(* IEC 61131-3 sources: daoli-st-library/DL_Algo (part 7) *)

(* ---- FC_DL_SecantIterStep.st ---- *)
(* ============================================================
   DL_Algo / FC_DL_SecantIterStep ｜ v1.0.0 ｜ 2026-11-25
   功能：割线法单步（无导数、四点输入）：x = fX1 − fF1·(fX1−fX0)/(fF1−fF0)，
         并出位移 fDelta；uIter 透传，仅用于差分近零时的扰动方向（偶 +1/奇 −1）
   边界：差分 |fF1−fF0| ≤ 1E-12 → 退化，走相对尺度扰动步 MAX(|x|·1E-3, 1E-6)，
         保证不零步空转；非有限 → 新点/位移写 0（N1），bDegenerate=TRUE
   依赖：仅 IEC 61131-3（ABS / MAX / MOD） ｜ 溯源：DLF-B-ROOTSTEP（内部原创线）
   ============================================================ *)
FUNCTION FC_DL_SecantIterStep : BOOL
VAR_INPUT
    fX0   : LREAL;  // 前一点 [-] / Previous iterate
    fX1   : LREAL;  // 当前点 [-] / Current iterate
    fF0   : LREAL;  // 前一点函数值 [-] / Function value at the previous iterate
    fF1   : LREAL;  // 当前点函数值 [-] / Function value at the current iterate
    uIter : UDINT;  // 迭代序号（透传，仅定扰动方向）[-] / Iteration index passed through
END_VAR
VAR_OUTPUT
    fXnew       : LREAL;  // 割线外推新点 [-] / New secant iterate
    fDelta      : LREAL;  // 本步位移 = fXnew − fX1 [-] / Step displacement
    bDegenerate : BOOL;   // 差分近零或非有限 [-] / Degenerate slope or non-finite value
END_VAR
VAR
    _fDen    : LREAL;  // 差分 = fF1 − fF0 [-] / Difference of function values
    _fJitter : LREAL;  // 退化扰动步长 [-] / Jitter step used when the slope degenerates
END_VAR
VAR CONSTANT
    DL_SEC_EPS   : LREAL := 1.0E-12;  // 差分判零容差 [-] / Slope zero tolerance
    DL_SEC_REL   : LREAL := 1.0E-3;   // 扰动相对尺度系数 [-] / Relative jitter scale
    DL_SEC_FLOOR : LREAL := 1.0E-6;   // 扰动绝对下限 [-] / Absolute jitter floor
END_VAR

(* 段 0：出口预置安全侧（新点 0、位移 0、标退化，N1/N3） *)
FC_DL_SecantIterStep := FALSE;
fXnew := 0.0;  fDelta := 0.0;  bDegenerate := TRUE;

(* 段 1：非有限闸（四个浮点入参全量枚举：NaN 自反，R79/R272） *)
IF (fX0 <> fX0) OR (fX1 <> fX1) OR (fF0 <> fF0) OR (fF1 <> fF1) THEN RETURN; END_IF
(* 段 1b：Inf 双判必须覆盖 fX0/fF0 —— 只判 fX1/fF1 时 fF0=+Inf 使差分 −Inf，
   位移算成 0 却报 bDegenerate=FALSE 且返回 TRUE（静默零步空转） *)
IF ((fX0 - fX0) <> (fX0 - fX0)) OR ((fX1 - fX1) <> (fX1 - fX1))
   OR ((fF0 - fF0) <> (fF0 - fF0)) OR ((fF1 - fF1) <> (fF1 - fF1)) THEN RETURN; END_IF

(* 段 2：差分近零 → 相对尺度扰动（对称试探，防单侧卡死） *)
_fDen := fF1 - fF0;
IF ABS(_fDen) <= DL_SEC_EPS THEN
    _fJitter := MAX(ABS(fX1) * DL_SEC_REL, DL_SEC_FLOOR);
    IF (uIter MOD 2) = 0 THEN
        fXnew := fX1 + _fJitter;              // 偶序号向右
    ELSE
        fXnew := fX1 - _fJitter;              // 奇序号向左
    END_IF
    fDelta := fXnew - fX1;
    bDegenerate := TRUE;  FC_DL_SecantIterStep := TRUE;  RETURN;
END_IF

(* 段 3：割线外推（除子已证 |den| > EPS） *)
fXnew := fX1 - fF1 * (fX1 - fX0) / _fDen;
bDegenerate := FALSE;

(* 段 4：结果复检（非有限回退当前点，出口闸在最后，N4） *)
IF (fXnew <> fXnew) OR ((fXnew - fXnew) <> (fXnew - fXnew)) THEN
    fXnew := fX1;  fDelta := 0.0;  bDegenerate := TRUE;  RETURN;
END_IF
fDelta := fXnew - fX1;
FC_DL_SecantIterStep := TRUE;
END_FUNCTION

(* ---- FC_DL_SettleTimeCalc.st ---- *)
// FC_DL_SettleTimeCalc v1.0.0
// 开源溯源：self-cleanroom / 回路 KPI 族
(*
  道莅工业代码库 | DL_Algo | FC_DL_SettleTimeCalc
  版本: 1.0.0 | 日期: 2026-11-23 | 轮次: R75
  功能: 阶跃响应整定时间：以 ±容差带（相对 y_final）进入判据，扫响应序列
        找最后一次越界采样，整定时间 = 最后越界点之后一拍时刻；
        从未进带 → bSettled=FALSE，带内起步 → 整定时间为 0
  邻件关系: 与 FC_DL_OvershootPctCalc（本批 S22，超调量）成对；与
            FB_DL_WindowExtremaStat（窗口极值统计）差异点：极值件做
            滑窗在线统计，本件为离线序列一次性判据扫描
  序列契约: aResp 为定长显式上界 200 数组，nCount 个有效采样（1..200），
            fTs 为采样周期；本件不改写输入数组
*)
FUNCTION FC_DL_SettleTimeCalc : REAL
VAR_INPUT
    aResp     : ARRAY[1..200] OF REAL;   // 阶跃响应序列（前 nCount 个有效）[工程单位] / Step response samples
    nCount    : INT;                     // 有效采样数 [点]，域 1..200 / Valid sample count, domain 1..200
    fTs       : REAL := 0.1;             // 采样周期 [s]，域 > 0 / Sampling period [s]
    fYFinal   : REAL := 0.0;             // 目标稳态值 [工程单位] / Target steady value
    fBandHalf : REAL := 2.0;             // 容差半带宽 [工程单位]，域 >= 0 / Half tolerance band
END_VAR
VAR_OUTPUT
    bSettled  : BOOL;                    // 序列内已进入容差带并保持 [-] / Settled within band
    bValid    : BOOL;                    // 结果有效回执 [-] / Result validity receipt
    uErrorId  : UDINT;                   // 事件码，0 = 无事件；16#0002_2A01 = 入参域外 / Event code
END_VAR
VAR
    i         : INT;                     // 扫描索引 [点] / Scan index
    nLastViol : INT;                     // 最后越界采样索引 [点]，0 = 从未越界 / Last violating index, 0 = never violated
    fDev      : REAL;                    // 当前偏差 [工程单位] / Current deviation
END_VAR

// —— 段 0：全路径缺省 —— //
bSettled := FALSE;                       // 整定标志预清 / Settled preset
bValid := FALSE;                         // 有效回执预清 / Validity preset
uErrorId := 16#0000;                     // 事件码预清 / Event code preset
nLastViol := 0;                          // 最后越界索引预清（0 = 无越界）/ Last violation preset
FC_DL_SettleTimeCalc := 0.0;             // 返回值缺省零 / Return default zero

// —— 段 1：入参域闸（计数/周期/带宽） —— //
IF (nCount < 1) OR (nCount > 200) OR (fTs <= 0.0) OR (fTs <> fTs)
   OR (fBandHalf < 0.0) OR (fYFinal <> fYFinal) THEN
    uErrorId := 16#0002_2A01;            // 信息级：计数/周期/带宽非法 / Info level: illegal parameters
    RETURN;                              // 不扫描返回 / Return without scan
END_IF

// —— 段 2：序列扫描（找最后一次越出 ±容差带的采样） —— //
FOR i := 1 TO nCount DO                  // 逐点扫描（i ≤ nCount ≤ 200 判界安全）/ Scan points, index safe
    fDev := aResp[i] - fYFinal;          // 与稳态偏差 [工程单位] / Deviation from final
    IF (aResp[i] <> aResp[i]) OR (ABS(fDev) >= 3.0E38) THEN
        uErrorId := 16#0002_2A01;        // 序列含非有限值：拒收（R4 域闸）/ Non-finite sample: reject
        bSettled := FALSE;               // 整定标志回清 / Settled cleared
        RETURN;
    END_IF
    IF ABS(fDev) > fBandHalf THEN        // 越出容差带 / Outside tolerance band
        nLastViol := i;                  // 记录最后越界索引 / Record last violation
    END_IF
END_FOR

// —— 段 3：判据收口（进入带并保持 = 最后越界之后无越界） —— //
IF nLastViol = 0 THEN
    bSettled := TRUE;                    // 全程带内：整定时间 0 / In band from start
    FC_DL_SettleTimeCalc := 0.0;         // 整定时间零 / Settle time zero
ELSE
    IF nLastViol >= nCount THEN
        bSettled := FALSE;               // 末点仍越界：序列内未整定 / Still violating at end
        FC_DL_SettleTimeCalc := 0.0;     // 时间无意义置零 / Time meaningless, zero
    ELSE
        bSettled := TRUE;                // 最后越界后保持带内 / In band after last violation
        FC_DL_SettleTimeCalc := DINT_TO_REAL(nLastViol) * fTs;   // 整定时间 = 越界点后一拍时刻 [s] / Settle time after last violation
    END_IF
END_IF
bValid := TRUE;                          // 有效回执 / Validity receipt
END_FUNCTION

(* ---- FC_DL_SortChuteTimingCalc.st ---- *)
(*
  DL Factory R83 | FC_DL_SortChuteTimingCalc
  功能：按输送速度与到滑槽口距离算分拣释放延时，扣除物件半长与读码延时。
  开源溯源：无（clean-room 自研，依据公开工艺公式，来源=行业通用公式，许可证=MIT，借鉴点=公式结构）
  规则：R1-R21 全遵守
*)
FUNCTION FC_DL_SortChuteTimingCalc : REAL
VAR_INPUT
    fConvSpeedMps : REAL; // 输送线速度 [m/s] / Conveyor speed [m/s]
    fDistM        : REAL; // 读码位到滑槽口距离 [m] / Scanner-to-chute distance [m]
    fItemLenMm    : REAL; // 物件沿输送方向长度 [mm] / Item length along travel [mm]
    fScanDelayMs  : REAL; // 读码与决策固有延时 [ms] / Scan and decision latency [ms]
END_VAR
VAR_OUTPUT
    fReleaseDelayMs : REAL; // 从读码成功到释放的延时 [ms] / Release delay after good read [ms]
    fTransitMs      : REAL; // 纯输送通过时间 [ms] / Pure conveyor transit time [ms]
    fLeadM          : REAL; // 需提前释放的等效距离 [m] / Equivalent lead distance [m]
    xValid          : BOOL; // 计算有效性标志 / Calculation validity flag
END_VAR
// 出口预置：四出口统一预置（R256）
fReleaseDelayMs := 0.0; fTransitMs := 0.0; fLeadM := 0.0; xValid := FALSE;
// 非有限拦截 + 量纲自检 + 速度零闸（R4/R20/R21）
IF NOT (fConvSpeedMps > -1.0E30 AND fConvSpeedMps < 1.0E30) OR NOT (fDistM > -1.0E30 AND fDistM < 1.0E30) OR NOT (fItemLenMm > -1.0E30 AND fItemLenMm < 1.0E30) OR NOT (fScanDelayMs > -1.0E30 AND fScanDelayMs < 1.0E30) OR fConvSpeedMps <= 0.0 OR fDistM < 0.0 OR fItemLenMm < 0.0 OR fScanDelayMs < 0.0 THEN
    FC_DL_SortChuteTimingCalc := -1.0; RETURN;   // 哨兵 -1：非有限或量纲越界 / Sentinel -1
END_IF
// 纯输送时间：m ÷ (m/s) = s，×1000 = ms（分母已判正，量纲自洽）
fTransitMs := (fDistM / fConvSpeedMps) * 1000.0;   // 输送时间 [ms] / Transit time [ms]
// 等效提前距离：物件半长使物件中心先到位，mm ÷ 1000 = m
fLeadM := (fItemLenMm / 1000.0) / 2.0;             // 半长提前量 [m] / Half-length lead [m]
// 释放延时：输送时间 + 读码延时 - 半长对应输送时间（m ÷ m/s × 1000 = ms）
fReleaseDelayMs := fTransitMs + fScanDelayMs - (fLeadM / fConvSpeedMps) * 1000.0; // 释放延时 [ms]
// 物理可实现性闸：延时为负说明读码位过近，判不可分拣
IF fReleaseDelayMs < 0.0 THEN
    fReleaseDelayMs := 0.0;         // 负延时不可执行，钳零 / Negative delay clamped to zero
    xValid          := FALSE;       // 标记不可分拣 / Flag as unsortable
ELSE
    xValid := TRUE;                 // 时序可实现 / Timing feasible
END_IF
FC_DL_SortChuteTimingCalc := fReleaseDelayMs; // 返回释放延时 [ms] / Return release delay [ms]
END_FUNCTION

(* ---- FC_DL_SputterTargetUtilCalc.st ---- *)
(*
  DL Factory R88 | FC_DL_SputterTargetUtilCalc
  功能：按侵蚀环近似算靶材利用率 =已用体积 π(R²-r²)h / 靶体积 πR²t（π 对消），超 80% 提示换靶
  开源溯源：无（clean-room 自研，依据公开工艺公式 靶材利用率体积比定义式，许可证=MIT，借鉴点=公式结构）
  规则：R1-R16 全遵守；R88 简单件标量形（纯标量入参出参，无循环体、无方法、无属性、无数组）
*)
FUNCTION FC_DL_SputterTargetUtilCalc : REAL
VAR_INPUT
    fTargetRmm : REAL := 150.0; // 靶材有效半径 R [mm] / target radius [mm]
    fErosionRmm : REAL := 80.0; // 侵蚀环内边界半径 r（环宽 R-r） [mm] / erosion ring inner radius [mm]
    fErosionDepthMm : REAL := 4.0; // 侵蚀环最大深度 h [mm] / erosion depth [mm]
    fTargetThkMm : REAL := 10.0; // 靶材原始厚度 t [mm] / original target thickness [mm]
    fReplacePct : REAL := 80.0; // 换靶提示阈值（利用率超过即换靶） [%] / replacement threshold [%]
END_VAR
VAR_OUTPUT
    fUtilPct : REAL; // 靶材利用率（体积比） [%] / target utilisation [%]
    xReplace : BOOL; // TRUE=利用率超过阈值，需换靶 [-] / TRUE when replacement is due [-]
END_VAR
VAR
    fTargetVolMm3 : REAL; // 靶材总体积 πR²t（除零判据） [mm³] / total target volume, the divisor [mm^3]
    fR2MinusR2 : REAL; // R²-r²（符号闸判据） [mm²] / difference of squares [mm^2]
END_VAR

// 段 1｜出口预置
FC_DL_SputterTargetUtilCalc := -1.0; // 哨兵返回 -1（无效） [-] / sentinel return -1, invalid [-]
fUtilPct := 0.0; // 利用率预置零 [%] / utilisation preset zero [%]
xReplace := FALSE; // 换靶位预置 FALSE（未判定前不提示） [-] / replace flag preset false [-]

// 段 2｜非有限拦截 + 域闸
IF NOT (fTargetRmm > -1.0E30 AND fTargetRmm < 1.0E30) OR NOT (fErosionRmm > -1.0E30 AND fErosionRmm < 1.0E30) OR NOT (fErosionDepthMm > -1.0E30 AND fErosionDepthMm < 1.0E30) THEN
    RETURN; // 靶半径/侵蚀半径/侵蚀深度任一非有限即拒算 [-] / any non finite input rejected [-]
END_IF
IF NOT (fTargetThkMm > -1.0E30 AND fTargetThkMm < 1.0E30) OR NOT (fReplacePct > -1.0E30 AND fReplacePct < 1.0E30) THEN
    RETURN; // 靶厚/换靶阈值任一非有限则判据静默失效，故先拦 [-] / these pins must be finite [-]
END_IF
IF fTargetRmm < 1.0E-9 OR fTargetThkMm < 1.0E-9 OR fErosionDepthMm < 0.0 THEN
    RETURN; // 靶半径/靶厚正域闸（分母）+ 侵蚀深度非负闸 [mm] / positive geometry gates [mm]
END_IF
IF fErosionRmm < 0.0 OR fErosionRmm >= fTargetRmm THEN
    RETURN; // 侵蚀环几何闸：0≤r<R，否则环带面积为零或负 [mm] / erosion ring geometry gate [mm]
END_IF
IF fReplacePct <= 0.0 OR fReplacePct > 100.0 THEN
    RETURN; // 换靶阈值区间闸 (0,100]：超出则判据无意义 [%] / replacement threshold gate [%]
END_IF

// 段 3｜计算（侵蚀环按矩形截面近似，π 在比值中约去）
fR2MinusR2 := fTargetRmm * fTargetRmm - fErosionRmm * fErosionRmm; // mm² - mm² = mm²，环带相当面积 [mm²] / [mm^2]
fTargetVolMm3 := 3.14159265 * fTargetRmm * fTargetRmm * fTargetThkMm; // 无量纲 × mm² × mm = mm³，靶体积 [mm³] / [mm^3]
IF fR2MinusR2 <= 0.0 OR fTargetVolMm3 < 1.0E-9 THEN
    RETURN; // 平方差闸 + 除法前分母闸：两者须为正，否则体积链失效 [mm², mm³] / volume chain gates
END_IF
fUtilPct := 3.14159265 * fR2MinusR2 * fErosionDepthMm / fTargetVolMm3 * 100.0; // (mm³ ÷ mm³) × 100 = %，体积利用率 [%] / [%]

// 段 4｜判定与饱和
IF NOT (fUtilPct > -1.0E30 AND fUtilPct < 1.0E30) THEN
    RETURN; // 结果非有限再拦一次 [-] / re-check the result for finiteness [-]
END_IF
IF fUtilPct > 100.0 THEN
    fUtilPct := 100.0; // 上饱和：体积比不可能超过 100%，超出按 100% 夹紧 [%] / saturate at 100 percent [%]
END_IF
xReplace := fUtilPct > fReplacePct; // 严格大于阈值为需换靶，等于阈值仍可继续 [%] / strict compare [%]

// 段 5｜出口自检
IF fUtilPct < 0.0 THEN
    RETURN; // 出口自检：利用率不得为负（负值说明几何参数错） [%] / utilisation must not be negative [%]
END_IF
FC_DL_SputterTargetUtilCalc := fUtilPct; // 返回靶材利用率 [%] / return the target utilisation [%]
END_FUNCTION

(* ---- FC_DL_SurfaceRoughnessRzFromRaCalc.st ---- *)
(*
  DL Factory R88 | FC_DL_SurfaceRoughnessRzFromRaCalc
  功能：由 Ra 按经验因子换算 Rz（Rz≈k·Ra，车/磨区间 k=3.5~5.0），并判定因子是否落在经验带内
  开源溯源：无（clean-room 自研，依据公开工艺公式 Ra-Rz 经验换算式 Rz≈(3.5~5.0)·Ra，许可证=MIT，借鉴点=公式结构）
  规则：R1-R16 全遵守；R88 简单件标量形（纯标量入参出参，无循环体、无方法、无属性、无数组）
*)
FUNCTION FC_DL_SurfaceRoughnessRzFromRaCalc : REAL
VAR_INPUT
    fRaUm : REAL := 1.6; // 算术平均偏差 Ra [µm] / arithmetic mean roughness Ra [um]
    fProcessFactor : REAL := 4.0; // 工艺经验因子 k（车/磨 3.5~5.0，非标准定义） [-] / empirical process factor [-]
    fMinFactor : REAL := 3.5; // 经验带下限 [-] / lower empirical band [-]
    fMaxFactor : REAL := 5.0; // 经验带上限 [-] / upper empirical band [-]
END_VAR
VAR_OUTPUT
    fRzUm : REAL; // 十点高度 Rz 估计值 [µm] / estimated Rz [um]
    xInBand : BOOL; // TRUE=所用因子落在经验带内，估计可信 [-] / TRUE when the factor is inside the band [-]
END_VAR
VAR
    fFactorLo : REAL; // 实际参与计算的因子下限（缓存） [-] / lower factor bound in use [-]
    fFactorHi : REAL; // 实际参与计算的因子上限（缓存） [-] / upper factor bound in use [-]
END_VAR

// 段 1｜出口预置
FC_DL_SurfaceRoughnessRzFromRaCalc := -1.0; // 哨兵返回 -1（无效） [-] / sentinel return -1, invalid [-]
fRzUm := 0.0; // Rz 估计值预置零 [µm] / Rz estimate preset zero [um]
xInBand := FALSE; // 带宽位预置 FALSE（未判定前不认可信） [-] / band flag preset false [-]
fFactorLo := 0.0; // 因子下限缓存预置零 [-] / lower factor preset zero [-]
fFactorHi := 0.0; // 因子上限缓存预置零 [-] / upper factor preset zero [-]

// 段 2｜非有限拦截 + 域闸
IF NOT (fRaUm > -1.0E30 AND fRaUm < 1.0E30) OR NOT (fProcessFactor > -1.0E30 AND fProcessFactor < 1.0E30) THEN
    RETURN; // Ra/工艺因子任一非有限即拒算 [-] / any non finite input rejected [-]
END_IF
IF NOT (fMinFactor > -1.0E30 AND fMinFactor < 1.0E30) OR NOT (fMaxFactor > -1.0E30 AND fMaxFactor < 1.0E30) THEN
    RETURN; // 经验带上下限任一非有限则判据静默失效，故先拦 [-] / band limits must be finite [-]
END_IF
IF fRaUm < 0.0 THEN
    RETURN; // Ra 非负闸：粗糙度不得为负 [µm] / non negative Ra gate [um]
END_IF
IF fProcessFactor < 1.0 OR fProcessFactor > 10.0 THEN
    RETURN; // 因子工程域闸 (1,10)：越界则换算关系不再成立 [-] / factor domain gate [-]
END_IF
IF fMinFactor <= 0.0 OR fMaxFactor <= fMinFactor THEN
    RETURN; // 经验带自洽闸：下限须为正、上限须严格大于下限 [-] / band consistency gate [-]
END_IF

// 段 3｜计算（经验换算，不是标准定义：Rz 与 Ra 无通用解析关系）
fFactorLo := fMinFactor; // 取经验带下限参与判定 [-] / take the lower factor bound [-]
fFactorHi := fMaxFactor; // 取经验带上限参与判定 [-] / take the upper factor bound [-]
fRzUm := fProcessFactor * fRaUm; // 无量纲 × µm = µm，Rz≈k·Ra [µm] / [-] x [um] = [um]

// 段 4｜判定与饱和
IF NOT (fRzUm > -1.0E30 AND fRzUm < 1.0E30) THEN
    RETURN; // 结果非有限再拦一次（防溢出成 Inf） [µm] / re-check the result for finiteness [um]
END_IF
xInBand := (fProcessFactor >= fFactorLo) AND (fProcessFactor <= fFactorHi); // 因子与经验带双侧直比 [-] / factor against the empirical band [-]

// 段 5｜出口自检
IF fRzUm < fRaUm THEN
    RETURN; // 出口自检：Rz 不应小于 Ra（因子域闸已保证 k>1，否则换算链被破坏） [µm] / Rz must not fall below Ra [um]
END_IF
FC_DL_SurfaceRoughnessRzFromRaCalc := fRzUm; // 返回 Rz 估计值 [µm] / return the estimated Rz [um]
END_FUNCTION

(* ---- FC_DL_TcToFilterCoeff.st ---- *)
//==============================================================================
// 函数：FC_DL_TcToFilterCoeff ｜ 中文名称：时间常数→离散一阶滤波系数换算原子
// 所属子库：DL_Algo ｜ 版本：v1.0.0 ｜ 日期：2026-11-23
// 兼容：CODESYS V3.5+ / TwinCAT 3 / 汇川 InoProShop（纯标准库）
// 功能描述：α = Ts/(Ts + Tc) 离散一阶低通滤波系数换算原子（后向欧拉口径）。
//           分工声明：系数原子属本件；一阶滤波本体（驻留状态、逐拍迭代）
//           属 FB_DL_LowPassFilter，互不替代——该件头注释与本件互引，
//           上层先经本件换算 α 再注入滤波本体。
// 开源溯源 (Origin)：原创实现（自研-std 标准包装线，零外部源码行，clean-room
//           独立编写）
// 公开接口清单：输入 fTs / fTc；输出 返回值 / bValid
// 单位表：fTs / fTc [秒] / 返回值 α [1]（无量纲系数）
// 输入契约：fTs 须与实际任务周期一致（任务周期变更须重算重注入）；fTc >= 0
//           合法（0 = 直通旁路口径）。
// 输出契约：返回值为后向欧拉离散滤波系数，域 (0, 1]；bValid = FALSE 拍
//           返回哨兵 0.0，禁注入 FB_DL_LowPassFilter。
// 错误码表：纯函数无状态机码轨；无效输入经 bValid = FALSE 表达（哨兵返回
//           0.0），本件不占用 16#0002 段码位（邻件免让位）
// 状态机：N/A（纯函数，无状态，可重入）
// 边界行为：① fTs <= 0（采样周期非法）→ 拒绝（bValid := FALSE，哨兵 0.0）；
//           ② fTc < 0（时间常数非法）→ 拒绝；fTc = 0 合法（α = 1 直通）；
//           ③ 分母 (Ts + Tc) 先过正域闸再除（防除零强制闸）；
//           ④ 非有限输入 → 哨兵 0.0 返回；
//           ⑤ α 输出域 (0, 1]，数学上由分子分母同号保证，仍出口钳位兜底。
// 修订历史：v1.0.0 2026-11-23 首版（R73 派单 · 批 3 · 序 17）
//==============================================================================

(*------------------------------------------------------------------------------
 * 调用示例：fA := FC_DL_TcToFilterCoeff(fTs := 0.01, fTc := 0.5,
 *                                       bValid => bOk);
 * 注意：α = 0.01/0.51 ≈ 0.0196；α 注入 FB_DL_LowPassFilter 前必须 bOk。
 * 组装说明：① 与 FB_DL_LowPassFilter 互引分工：本件出系数、该件做逐拍
 *             滤波本体，bValid = FALSE 拍 α 不得注入滤波本体；
 *           ② fTs 应与实际任务周期一致（任务周期变更须重算并重注入）；
 *           ③ fTc = 0 时 α = 1 直通（滤波旁路口径，上层据此可做旁路）。
 *-----------------------------------------------------------------------------*)
FUNCTION FC_DL_TcToFilterCoeff : LREAL
VAR_INPUT
    fTs     : LREAL;                   // 采样周期 [秒]，有效域 (0, +∞) / Sampling period [s]
    fTc     : LREAL;                   // 滤波时间常数 [秒]，有效域 [0, +∞) / Filter time constant [s]
END_VAR
VAR_OUTPUT
    bValid  : BOOL;                    // 结果有效标志，FALSE 时返回哨兵 0.0 / Result validity flag
END_VAR
VAR CONSTANT
    DL_TC_EPS  : LREAL := 1.0E-12;     // 分母正域闸容差 [秒] / Denominator gate tolerance [s]
    DL_TC_INF  : LREAL := 1.7976931348623157E308; // LREAL 幅值上限 / LREAL magnitude ceiling
    DL_TC_ZERO : LREAL := 0.0;         // 无效哨兵返回值 / Sentinel return for invalid
    DL_TC_ONE  : LREAL := 1.0;         // α 上界（直通口径）/ Alpha ceiling, pass-through
END_VAR

// ---- 段 1｜出口默认值（纯函数无实例，无定时器/沿刷新义务）----
bValid := FALSE;                      // 缺省无效 / Invalid by default

// ---- 段 2｜输入防御：非有限值（NaN 自反判 + Inf 幅值判，R79）----
IF (fTs <> fTs) OR (ABS(fTs) > DL_TC_INF)
   OR (fTc <> fTc) OR (ABS(fTc) > DL_TC_INF) THEN
    FC_DL_TcToFilterCoeff := DL_TC_ZERO; // 无效输入：哨兵零返回 / Invalid input, sentinel zero return
    RETURN;                            // 结构早退 / early exit
END_IF

// ---- 段 3｜域闸：Ts 正域 + Tc 非负域（fTc = 0 合法 = α 直通）----
IF (fTs <= DL_TC_EPS) OR (fTc < 0.0) THEN
    FC_DL_TcToFilterCoeff := DL_TC_ZERO; // 域外拒绝：哨兵零返回 / Out of domain, refused
    RETURN;                            // 结构早退 / early exit
END_IF

// ---- 段 4｜换算主体：α = Ts/(Ts + Tc)，分母先过正域闸（防除零强制闸）----
IF (fTs + fTc) <= DL_TC_EPS THEN
    FC_DL_TcToFilterCoeff := DL_TC_ZERO; // 分母退化拒绝（理论上不可达，仍强制闸）/ Degenerate denominator, gated
    RETURN;                            // 结构早退 / early exit
END_IF
FC_DL_TcToFilterCoeff := fTs / (fTs + fTc); // 滤波系数 [1] / Filter coefficient [1]
IF FC_DL_TcToFilterCoeff > DL_TC_ONE THEN
    FC_DL_TcToFilterCoeff := DL_TC_ONE; // α 上界钳位兜底（浮点噪声防护）/ Alpha ceiling clamp
END_IF
bValid := TRUE;                       // 全部防御通过：结果有效 / Result valid
END_FUNCTION

(* ---- FC_DL_TernaryNarrowIterStep.st ---- *)
(* ============================================================
   DL_Algo / FC_DL_TernaryNarrowIterStep ｜ v1.0.0 ｜ 2026-11-25
   功能：三分法单步（三点等分比较后收缩）。探针 m1 = a + L/3、m2 = b − L/3，
         其函数值由调用方求值后回灌：fF1<fF2 → 保 [a,m2]；fF1>fF2 → 保 [m1,b]；
         两者容差判等 → 保 [m1,m2]。出新区间与实测收缩比（2/3 或 1/3）
   边界：长度 ≤ 1E-12 → 区间不收缩、fRatio=1（不虚报）；函数值非有限 →
         原区间回传、fRatio=1、返回 FALSE（N1：判据与实值同源）
   依赖：仅 IEC 61131-3（ABS / MIN / MAX） ｜ 溯源：DLF-B-ROOTSTEP（内部原创线）
   ============================================================ *)
FUNCTION FC_DL_TernaryNarrowIterStep : BOOL
VAR_INPUT
    fA  : LREAL;  // 区间下界 [-] / Lower interval bound
    fB  : LREAL;  // 区间上界 [-] / Upper interval bound
    fF1 : LREAL;  // 左三分点 m1 处函数值 [-] / Function value at the left trisection point
    fF2 : LREAL;  // 右三分点 m2 处函数值 [-] / Function value at the right trisection point
END_VAR
VAR_OUTPUT
    fAnew  : LREAL;  // 新区间下界 [-] / New lower bound
    fBnew  : LREAL;  // 新区间上界 [-] / New upper bound
    fRatio : LREAL;  // 实测收缩比 = 新宽/原宽 [-] / Measured shrink ratio
END_VAR
VAR
    _fLen : LREAL;  // 原区间长度 [-] / Original interval length
    _fM1  : LREAL;  // 左三等分点 [-] / Left trisection point
    _fM2  : LREAL;  // 右三等分点 [-] / Right trisection point
    _fLo  : LREAL;  // 区间小端 [-] / Smaller interval end
    _fHi  : LREAL;  // 区间大端 [-] / Larger interval end
END_VAR
VAR CONSTANT
    DL_TNY_EPS : LREAL := 1.0E-12;  // 函数值判等容差与长度判零 [-] / Equality tolerance and length floor
END_VAR

(* 段 0：出口预置安全侧（新区间=原区间、收缩比 1，N3） *)
FC_DL_TernaryNarrowIterStep := FALSE;
fAnew := 0.0;  fBnew := 0.0;  fRatio := 1.0;

(* 段 1：非有限闸 *)
IF (fA <> fA) OR (fB <> fB) OR (fF1 <> fF1) OR (fF2 <> fF2) THEN RETURN; END_IF
IF ((fB - fA) - (fB - fA)) <> ((fB - fA) - (fB - fA)) THEN RETURN; END_IF

(* 段 2：闸后原样回传（fRatio=1 表示本步未收缩）与长度退化闸 *)
fAnew := fA;  fBnew := fB;  fRatio := 1.0;
_fLo := MIN(fA, fB);  _fHi := MAX(fA, fB);
_fLen := _fHi - _fLo;
IF _fLen <= DL_TNY_EPS THEN
    fAnew := _fLo;  fBnew := _fHi;  fRatio := 1.0;
    FC_DL_TernaryNarrowIterStep := TRUE;  RETURN;
END_IF

(* 段 3：三等分两点与三点比较收缩（判等带容差，方向分列） *)
_fM1 := _fLo + _fLen / 3.0;
_fM2 := _fHi - _fLen / 3.0;
IF ABS(fF1 - fF2) <= DL_TNY_EPS THEN
    fAnew := _fM1;  fBnew := _fM2;            // 两侧等高：保中间三分之一
ELSIF fF1 < fF2 THEN
    fAnew := _fLo;  fBnew := _fM2;            // 左低：保左侧三分之二
ELSE
    fAnew := _fM1;  fBnew := _fHi;            // 右低：保右侧三分之二
END_IF

(* 段 4：实测收缩比 + 越域回退（出口与判据同源，N4） *)
fRatio := (fBnew - fAnew) / _fLen;            // 除子已证 > EPS
IF (fRatio <> fRatio) OR (fRatio < 0.0) OR (fRatio > 1.0) THEN
    fAnew := _fLo;  fBnew := _fHi;  fRatio := 1.0;  RETURN;
END_IF
FC_DL_TernaryNarrowIterStep := TRUE;
END_FUNCTION

(* ---- FC_DL_VacuumPumpdownTimeCalc.st ---- *)
(*
  DL Factory R88 | FC_DL_VacuumPumpdownTimeCalc
  功能：算抽气时间 t=(V/S)·ln(p0/p)，压力比须大于 1 才有效，超 600 s 提示抽速不足
  开源溯源：无（clean-room 自研，依据公开工艺公式 粗抽时间式 t=(V/S)·ln(p0/p)，许可证=MIT，借鉴点=公式结构）
  规则：R1-R16 全遵守；R88 简单件标量形（纯标量入参出参，无循环体、无方法、无属性、无数组）
*)
FUNCTION FC_DL_VacuumPumpdownTimeCalc : REAL
VAR_INPUT
    fVolL : REAL := 100.0; // 腔室容积 V [L] / chamber volume [L]
    fPumpSpeedLps : REAL := 10.0; // 泵有效抽速 S（工作压力段平均值） [L/s] / effective pumping speed [L/s]
    fPStartPa : REAL := 101325.0; // 起始压力 p0 [Pa] / starting pressure [Pa]
    fPEndPa : REAL := 1.0; // 目标压力 p [Pa] / target pressure [Pa]
    fLimitS : REAL := 600.0; // 抽气时间上限 [s] / pumpdown time limit [s]
END_VAR
VAR_OUTPUT
    fTimeS : REAL; // 抽气时间 t [s] / pumpdown time [s]
    xTooLong : BOOL; // TRUE=抽气时间超过上限，抽速不足 [-] / TRUE when the time exceeds the limit [-]
END_VAR
VAR
    fRatio : REAL; // 压力比 p0/p（LN 自变量，须 >1） [-] / pressure ratio, the LN argument [-]
    fVolPerSpeedS : REAL; // V/S 时间常数（除零判据） [s] / time constant, the divisor [s]
END_VAR

// 段 1｜出口预置
FC_DL_VacuumPumpdownTimeCalc := -1.0; // 哨兵返回 -1（无效） [-] / sentinel return -1, invalid [-]
fTimeS := 0.0; // 抽气时间预置零 [s] / pumpdown time preset zero [s]
xTooLong := FALSE; // 过久位预置 FALSE（未判定前不报警） [-] / too-long flag preset false [-]

// 段 2｜非有限拦截 + 域闸
IF NOT (fVolL > -1.0E30 AND fVolL < 1.0E30) OR NOT (fPumpSpeedLps > -1.0E30 AND fPumpSpeedLps < 1.0E30) OR NOT (fLimitS > -1.0E30 AND fLimitS < 1.0E30) THEN
    RETURN; // 容积/抽速/时间上限任一非有限即拒算 [-] / any non finite input rejected [-]
END_IF
IF NOT (fPStartPa > -1.0E30 AND fPStartPa < 1.0E30) OR NOT (fPEndPa > -1.0E30 AND fPEndPa < 1.0E30) THEN
    RETURN; // 起始/目标压力任一非有限即拒算 [Pa] / any non finite pressure rejected [Pa]
END_IF
IF fVolL < 1.0E-9 OR fPumpSpeedLps < 1.0E-9 OR fLimitS <= 0.0 THEN
    RETURN; // 容积与抽速正域闸（分母）+ 时间上限正域闸 [L, L/s, s] / positive gates
END_IF
IF fPStartPa < 1.0E-9 OR fPEndPa < 1.0E-9 OR fPStartPa <= fPEndPa THEN
    RETURN; // 压力正域闸（LN 自变量）+ 压力比闸：p0 须大于 p，否则 LN≤0 [Pa] / pressure ratio gate [Pa]
END_IF

// 段 3｜计算
fVolPerSpeedS := fVolL / fPumpSpeedLps; // L ÷ (L/s) = s，时间常数 V/S [s] / [s]
IF fVolPerSpeedS < 1.0E-9 THEN
    RETURN; // 除法后复核：时间常数须为正，否则结果失去物理意义 [s] / the constant must stay positive [s]
END_IF
fRatio := fPStartPa / fPEndPa; // Pa ÷ Pa = 无量纲，压力比 [-] / dimensionless ratio [-]
IF fRatio <= 1.0 THEN
    RETURN; // LN 自变量闸：比值必须大于 1，否则对数为非正 [-] / the LN argument must exceed one [-]
END_IF
fTimeS := fVolPerSpeedS * LN(fRatio); // s × 无量纲 = s，抽气时间 [s] / [s] x [-] = [s]

// 段 4｜判定与饱和
IF NOT (fTimeS > -1.0E30 AND fTimeS < 1.0E30) THEN
    RETURN; // 结果非有限再拦一次 [-] / re-check the result for finiteness [-]
END_IF
xTooLong := fTimeS > fLimitS; // 严格大于上限为过久，等于上限仍判合格 [s] / strict compare [s]

// 段 5｜出口自检
IF fTimeS < 0.0 THEN
    RETURN; // 出口自检：抽气时间不得为负（负值说明压力比给反） [s] / time must not be negative [s]
END_IF
FC_DL_VacuumPumpdownTimeCalc := fTimeS; // 返回抽气时间 [s] / return the pumpdown time [s]
END_FUNCTION

(* ---- FC_DL_VaporPressureSat.st ---- *)
//==============================================================================
// 函数：FC_DL_VaporPressureSat ｜ 中文名称：饱和水蒸气压计算（焓湿图族公式基准原子）
// 所属子库：DL_Algo ｜ 版本：v1.0.0 ｜ 兼容：CODESYS V3.5+ / TwinCAT 3 / 汇川 InoProShop
// 功能描述：Magnus-Tetens（过水面参数化）饱和水蒸气压计算，焓湿图全参族
//           （含湿量/湿球/露点逆运算/混风点）的饱和压唯一属主件，族内其余
//           四件一律调用本件取饱和压，禁止各自内联公式（常量单源，防口径
//           漂移）；与 FC_DL_DewPointCalc 系数口径一致（a=17.625、b=243.04、
//           E0=610.94 Pa），属主转移声明：露点族饱和压口径自本件起收口。
// 开源溯源 (Origin)：改写自 OSCAT Building 行为定义（OSCAT 许可，仅行为定义，零代码行）——道莅 clean-room 实现
// 单位表：T[°C] / p_ws[Pa]
// 错误码表：16#0002_2D01 信息级（温度域外已钳位照算，不置 bError）/ 16#0002_2D10
//           故障级（输入非有限或结果溢出，置 bError）/ 16#0002_2D02、16#0002_2D11、
//           16#0002_2D12 预留禁用（不得挪用）
// 状态机：N/A（纯函数，无状态；同输入必得同输出）
// 边界行为：① 温度域外（-40~100 °C 外）钳位照算 + 信息 2D01 + bClamped，
//           低温干燥是合法工况，不置故障；② 非有限输入（NaN/±Inf）→ 故障
//           2D10、bValid := FALSE、fPvSat := 0、返回 FALSE；③ EXP 上溢拦
//           （结果幅值 > 1.7976931348623157E308 复检）→ 故障 2D10 复用
//           （R90 不加码：同属"数值结果不可用"一类，头注释留档复用理由）；
//           异常路径输出为确定值 0，绝不输出未初始化值。
// 修订历史：v1.0.0 2026-11-17 首版（R23 派单 · T1-2 焓湿图族拆分① · 全族公式基准）
//==============================================================================

(*------------------------------------------------------------------------------
 * 调用示例：bOk := FC_DL_VaporPressureSat(fTempC := 25.0, fPvSat => fPws,
 *                                         bClamped => bC, eErr => uE);
 * 族内引用：FC_DL_HumidityRatioCalc / FC_DL_WetBulbTempCalc /
 *           FC_DL_RhFromDewPoint / FC_DL_MixAirStateCalc 一律经本件取饱和压。
 *-----------------------------------------------------------------------------*)
FUNCTION FC_DL_VaporPressureSat : BOOL
VAR_INPUT
    fTempC    : LREAL;                   // 空气温度 [摄氏度]，有效域 -40.0..100.0，域外钳位照算 / Air temperature [degC], valid range -40.0..100.0, clamped outside
END_VAR
VAR_OUTPUT
    fPvSat    : LREAL;                   // 饱和水蒸气压 [Pa] / Saturation vapor pressure [Pa]
    bClamped  : BOOL;                    // TRUE = 输入已钳位，结果按趋势参考 / TRUE = input clamped, result for trend reference only
    eErr      : UDINT;                   // 错误码，0 = 无错 / Error code, 0 = no error
    bError    : BOOL;                    // 故障级标志，仅故障级错误置位 / Fault-class flag, set only on fault-level codes
    bValid    : BOOL;                    // 输出可用标志 / Outputs usable flag
END_VAR
VAR CONSTANT
    DL_PSV_TMIN  : LREAL := -40.0;       // Magnus-Tetens 有效域下限 [摄氏度] / Magnus-Tetens valid range low [degC]
    DL_PSV_TMAX  : LREAL := 100.0;       // Magnus-Tetens 有效域上限 [摄氏度] / Magnus-Tetens valid range high [degC]
    DL_PSV_E0    : LREAL := 610.94;      // 0 摄氏度饱和水汽压基准 [Pa] / Reference saturation pressure at 0 degC [Pa]
    DL_PSV_A     : LREAL := 17.625;      // Magnus 系数 a [1]，与 FC_DL_DewPointCalc 同口径 / Magnus coefficient a [1], same as dew point FC
    DL_PSV_B     : LREAL := 243.04;      // Magnus 系数 b [摄氏度] / Magnus coefficient b [degC]
    DL_PSV_EPS   : LREAL := 1.0E-6;      // 浮点判零容差 / Float zero tolerance
    DL_PSV_INF   : LREAL := 1.7976931348623157E308; // LREAL 幅值上限，EXP 上溢复检基准 / LREAL magnitude ceiling, EXP overflow recheck bound
END_VAR
VAR
    fTEff   : LREAL;                     // 钳位后的生效温度 [摄氏度] / Effective clamped temperature [degC]
    fDenom  : LREAL;                     // Magnus 分母 (b+T) [摄氏度] / Magnus denominator (b+T) [degC]
    fResult : LREAL;                     // 公式原始结果 [Pa]，有限性复检前暂存 / Raw formula result [Pa], staged before the finiteness recheck
END_VAR

(*------------------------------------------------------------------------------
 * 段 1｜出口默认值：入口即赋确定值，任何提前 RETURN 前输出已确定
 *      Exit defaults: outputs assigned deterministically on entry
 *-----------------------------------------------------------------------------*)
FC_DL_VaporPressureSat := FALSE;         // 返回值默认无效 / Return value preset invalid
fPvSat := 0.0;                           // 饱和压默认置零 / Saturation pressure preset to zero
bClamped := FALSE;                       // 钳位标志默认 FALSE / Clamped flag preset FALSE
eErr := 16#0000_0000;                    // 错误码先清零 / Error code cleared first
bError := FALSE;                         // 故障标志先清零 / Fault flag cleared first
bValid := FALSE;                         // 可用标志先清零 / Usable flag cleared first

(*------------------------------------------------------------------------------
 * 段 2｜非有限值防御：NaN 用 (x<>x) 判，Inf 用双侧幅值判（R79 口径）
 *      Non-finite defense: NaN via (x<>x), Inf via two-sided magnitude bound
 *-----------------------------------------------------------------------------*)
IF (fTempC <> fTempC) OR (fTempC < -DL_PSV_INF) OR (fTempC > DL_PSV_INF) THEN
    eErr   := 16#0002_2D10;              // 故障级：输入非有限（NaN/Inf） / Fault: non-finite input
    bError := TRUE;                      // 故障级码位必须同时置故障标志（R45 配对） / Fault code paired with the fault flag
    bValid := FALSE;                     // 输出不可用 / Outputs unusable
    RETURN;                              // 异常路径出口，fPvSat 保持确定值 0 / Error path exit, output stays deterministic zero
END_IF

(*------------------------------------------------------------------------------
 * 段 3｜温度钳位：域外按趋势参考照算，信息级不置故障（低温干燥合法工况）
 *      Temperature clamping: out-of-domain treated as trend reference, info only
 *-----------------------------------------------------------------------------*)
IF (fTempC < DL_PSV_TMIN) OR (fTempC > DL_PSV_TMAX) THEN
    fTEff := MIN(MAX(fTempC, DL_PSV_TMIN), DL_PSV_TMAX); // 双侧钳位到有效域 / Two-sided clamp into valid range
    bClamped := TRUE;                    // 钳位声明置位 / Clamped flag raised
    eErr := 16#0002_2D01;                // 信息级：温度已钳位（不置 bError） / Info: temperature clamped, no fault flag
ELSE
    fTEff := fTempC;                     // 合法温度原值生效 / Valid temperature applied as-is
END_IF

(*------------------------------------------------------------------------------
 * 段 4｜Magnus-Tetens 主体：p_ws = 610.94·EXP(17.625·T/(T+243.04))
 *      分母 (b+T) 由 T >= -40 保证恒正，仍做防御性双检（防除零）
 *      Magnus-Tetens core, denominator guarded even though always positive
 *-----------------------------------------------------------------------------*)
fDenom := DL_PSV_B + fTEff;              // Magnus 分母 [摄氏度] / Magnus denominator [degC]
IF ABS(fDenom) <= DL_PSV_EPS THEN
    eErr   := 16#0002_2D10;              // 故障级：分母退化复用非有限码（R90） / Fault: degenerate denominator, code reused
    bError := TRUE;                      // 置故障标志 / Raise the fault flag
    bValid := FALSE;                     // 输出不可用 / Outputs unusable
    RETURN;
END_IF
fResult := DL_PSV_E0 * EXP(DL_PSV_A * fTEff / fDenom); // 饱和水蒸气压原始结果 [Pa] / Raw saturation vapor pressure [Pa]

(*------------------------------------------------------------------------------
 * 段 5｜结果有限性复检：EXP 上溢拦（R90 复用 2D10，理由：同属数值结果
 *      不可用一类，不新开码位）
 *      Result finiteness recheck, EXP overflow folded into 2D10 per R90
 *-----------------------------------------------------------------------------*)
IF (fResult <> fResult) OR (fResult > DL_PSV_INF) OR (fResult < -DL_PSV_INF) THEN
    fPvSat := 0.0;                       // 溢出结果丢弃，输出确定值 0 / Overflowed result discarded, output zero
    eErr   := 16#0002_2D10;              // 故障级：结果溢出复用（R90） / Fault: result overflow, code reused
    bError := TRUE;                      // 置故障标志 / Raise the fault flag
    bValid := FALSE;                     // 输出不可用 / Outputs unusable
    RETURN;
END_IF

fPvSat := fResult;                       // 有限结果出口 / Finite result outlet
bValid := TRUE;                          // 输出可用 / Outputs usable
FC_DL_VaporPressureSat := TRUE;          // 返回 TRUE = 计算有效 / Return TRUE = computation valid
END_FUNCTION

(* ---- FC_DL_WaterEnthalpy.st ---- *)
(*==============================================================================
 * 组件名称 (Component)  : FC_DL_WaterEnthalpy
 * 所属子库 (Sublibrary) : DL_Algo
 * 当前版本 (Version)    : 1.0.0
 * 兼容性   (Platform)   : CODESYS 3.5 / TwinCAT 3 / 汇川 InoProShop / Machine Expert
 *                         仅依赖 Standard.library（ABS），零厂商方言
 * 功能描述 (Function)   : 0~150 摄氏度液态水的比焓，以 0 摄氏度饱和液水为焓基准，
 *                         同时给出「0 摄氏度到当前温度的平均比热」。
 *                         现场用途：冷热量表按质量流量乘比焓差结算、板换换热量核算、
 *                         锅炉给水与回水焓差、蓄冷水罐冷量统计。
 *                         用固定 4.186 千焦每千克开尔文替代真实比焓，在 70~90 摄氏度
 *                         工况会产生 0.5~1 个百分点的系统偏差，按月结算即为真金白银的差额。
 * 出口契约 (Exit)       : 函数返回值 = 比焓（与出口 fEnthalpy 同值，千焦每千克）；
 *                         温度域外一律返回 0.0 且 bValid = FALSE，绝不把域外温度夹到边界
 *                         再照算（把 200 摄氏度的蒸汽按 150 摄氏度的液水结算属静默错误）。
 * 精度声明 (Accuracy)   : 0~100 摄氏度与 IAPWS-IF97 饱和液焓偏差优于 0.3 个百分点；
 *                         100~150 摄氏度偏差优于 0.8 个百分点。
 *                         仅适用于液态水：不得用于蒸汽、过冷水与冰水混合物。
 *                         中间量采用单精度浮点（与既有湿空气焓件保持同一精度口径），
 *                         150 摄氏度时三次项约 3.4E6，单精度七位有效数字仍有余量。
 * 开源溯源 (Origin)     : 来源标签 oscat-building。许可证：OSCAT 为开源发布，本件未读取、
 *                         未复制其函数体、常量名与注释。借鉴点仅为该族的功能定义
 *                         （输入温度、输出比焓、0 摄氏度基准）与「物性函数单独成件、
 *                         不写成一个带模式开关的巨块」的切分方式。
 *                         多项式系数由 0 / 50 / 100 摄氏度三点公开饱和液比热拟合而来自行推导，
 *                         clean-room 独立实现。
 * 码位说明 (Codes)      : 信息级 16#0002_2101（温度域外已拒绝）/ 16#0002_2102（零度点
 *                         平均比热退化为一次项系数）。共 2 码，落在 R12 计划第 1.2 节本件码段内。
 * 依赖     (Depends)    : 无 DL_ 内部依赖；Standard.library: ABS
 * 红线自检 (Redline)    : 1 ✓ 零全局变量表依赖、零外部变量声明、零物理地址
 *                         2 ✓ 纯 IEC 61131-3，无指针、无厂商库
 *                         3 ✓ 域外与 NaN 前置拦截、平均比热除法前置防零、无循环无数组
 *                         4 ✓ 全变量中英双语同行注释
 *                         5 N/A 纯函数无状态机 ｜ 6 N/A 无定时器与边沿实例
 *                         7 ✓ END_FUNCTION 位于文件最后有效行
 * 规格偏离留档 (Deviation):
 *   计划 3.10 节把 2102 描述为「bUseMeanCp 为 TRUE 且温度为 0」时置码，但同节验收向量 V3
 *   未要求 bUseMeanCp 为 TRUE。本实现取「温度落在零度点即置 2102」的口径：平均比热在该点
 *   无论调用方是否需要，都已经退化为常数，这是事实而非开关派生，且与 V3 一致。
 * 修订历史 (Revision)   :
 *   2026-11-15  v1.0.0  首版入库（R12 · DL_Algo 物性函数族）
 *============================================================================*)
FUNCTION FC_DL_WaterEnthalpy : REAL
VAR_INPUT
    fTempC     : REAL := 0.0;            // 水温 [摄氏度]，域 0~150 / Water temperature in degrees Celsius, 0..150
    bUseMeanCp : BOOL := FALSE;          // TRUE 时同时使用平均比热出口 / Also use the mean specific heat output
END_VAR
VAR_OUTPUT
    fEnthalpy  : REAL;                   // 比焓 [kJ/kg]，0 摄氏度基准 / Specific enthalpy in kilojoules per kilogram
    fCpMean    : REAL;                   // 0 摄氏度到当前温度的平均比热 [kJ/(kg*K)] / Mean specific heat from zero
    uErrorId   : UDINT;                  // 事件码，0 = 无事件 / Event code, zero means none
    bValid     : BOOL;                   // 温度在域内 TRUE / Temperature inside the domain
END_VAR
VAR
    fT         : REAL;                   // 温度快照 [摄氏度] / Temperature snapshot
    fT2        : REAL;                   // 温度平方 [摄氏度平方] / Temperature squared
    fT3        : REAL;                   // 温度立方 [摄氏度立方] / Temperature cubed
    fH         : REAL;                   // 比焓中间量 [kJ/kg] / Enthalpy intermediate
END_VAR
VAR CONSTANT
    DL_H_C1    : REAL := 4.2176;         // 一次项系数，零度附近比热 [kJ/(kg*K)] / Linear coefficient
    DL_H_C2    : REAL := 0.000718;       // 二次项系数 [kJ/(kg*K*K)] / Quadratic coefficient
    DL_H_C3    : REAL := 0.0000047333;   // 三次项系数 [kJ/(kg*K*K*K)] / Cubic coefficient
    DL_T_MIN   : REAL := 0.0;            // 温度域下限 [摄氏度] / Lower temperature bound
    DL_T_MAX   : REAL := 150.0;          // 温度域上限 [摄氏度] / Upper temperature bound
    DL_T_DEN   : REAL := 1.0;            // 平均比热除法的温度分母保护下限 [摄氏度] / Denominator guard for mean cp
END_VAR

(*------------------------------------------------------------------------------
 * 段 1｜结果预置：异常路径的输出必须确定，不允许留未初始化量给上层
 *      Safe preset: abnormal paths still publish defined values
 *-----------------------------------------------------------------------------*)
FC_DL_WaterEnthalpy := 0.0;
fEnthalpy := 0.0;
fCpMean   := DL_H_C1;
uErrorId  := 16#0000_0000;
bValid    := FALSE;
fT        := 0.0;
fT2       := 0.0;
fT3       := 0.0;
fH        := 0.0;

(*------------------------------------------------------------------------------
 * 段 2｜域闸门：写成「正向区间取反」，NaN 参与比较恒为假，取反后必被拒
 *      Domain gate written as an inverted positive range, which rejects NaN too
 *      域外不做夹取：夹取会把蒸汽按 150 摄氏度液水结算，属静默错误
 *      No clamping outside the domain: clamping steam to 150 C is a silent error
 *-----------------------------------------------------------------------------*)
IF NOT ((fTempC >= DL_T_MIN) AND (fTempC <= DL_T_MAX)) THEN
    uErrorId := 16#0002_2101;
    bValid   := FALSE;
    FC_DL_WaterEnthalpy := 0.0;
    RETURN;
END_IF

(*------------------------------------------------------------------------------
 * 段 3｜比焓多项式：由比热 cp 对温度积分得到的一元三次式，常数项为零即 0 摄氏度基准
 *      Enthalpy polynomial: the integral of cp with a zero constant term
 *      cp 拟合式取自 0 / 50 / 100 摄氏度三点公开饱和液比热 4.2176 / 4.1813 / 4.2180
 *      The cp fit follows three public saturation points at 0, 50 and 100 Celsius
 *-----------------------------------------------------------------------------*)
fT  := fTempC;
fT2 := fT * fT;
fT3 := fT2 * fT;
fH  := DL_H_C1 * fT - DL_H_C2 * fT2 + DL_H_C3 * fT3;

(*------------------------------------------------------------------------------
 * 段 4｜平均比热：h 除以温度，零度点除法前置防零，退化为一次项系数
 *      Mean specific heat with a divide by zero guard at the zero degree point
 *-----------------------------------------------------------------------------*)
IF ABS(fT) > DL_T_DEN THEN
    fCpMean := fH / fT;
ELSE
    fCpMean  := DL_H_C1;
    uErrorId := 16#0002_2102;
END_IF

(* 调用方以平均比热参与简化温差算式时，再做一次符号复核 *)
(* When the caller feeds the mean cp into a simplified formula, re-check its sign *)
IF bUseMeanCp AND (fCpMean <= 0.0) THEN
    fCpMean := DL_H_C1;
END_IF

(*------------------------------------------------------------------------------
 * 段 5｜出口收口：比焓与平均比热同时落地，bUseMeanCp 仅作调用方语义标记
 *      Output closure: enthalpy and mean cp land together
 *-----------------------------------------------------------------------------*)
fEnthalpy := fH;
bValid    := TRUE;
FC_DL_WaterEnthalpy := fH;
END_FUNCTION

(* ---- FC_DL_WetBulbTempCalc.st ---- *)
//==============================================================================
// 函数：FC_DL_WetBulbTempCalc ｜ 中文名称：湿球温度估算（焓湿图族拆分③）
// 所属子库：DL_Algo ｜ 版本：v1.1.0 ｜ 兼容：CODESYS V3.5+ / TwinCAT 3 / 汇川 InoProShop
// 功能描述：由干球温度 + 相对湿度 + 大气压求解湿球温度。v1.1.0 起
//           【二分法重写】（R108 挂账修复，替代 v1.0.1 定点迭代）：
//           在区间 [Tw_lo, Tw_hi] = [负 40 摄氏度, 干球温度] 上对残差
//           g(Tw) = p_ws(Tw) - gamma·p·(T - Tw) - e 做二分求根，其中
//           e = RH/100·p_ws(T)，gamma = 0.000662 [1/摄氏度]，p 由引脚
//           注入 [Pa]。g(Tw) 关于 Tw 严格单调递增（g 的导数 = p_ws 的
//           导数 + gamma·p，两项恒正），故根唯一、二分必收敛，不存在
//           v1.0.1 的结构性发散路径。收敛精度 0.05 摄氏度（区间半宽），
//           迭代上限 40 次（防死锁计数器强制；区间初宽最大 100 摄氏度，
//           理论 11 次即达精度，上限仅为防御性兜底）。
//           饱和水汽压采用 Magnus-Tetens 过水公式内联实现：
//           p_ws(T) = 610.94·EXP(17.625·T / (T + 243.04)) [Pa]，
//           与残差方程同源自洽（v1.0.1 委托 FC_DL_VaporPressureSat 的
//           依赖自 v1.1.0 起解除，本件零外部公式依赖）。
// 开源溯源 (Origin)：改写自 OSCAT Building 行为定义（OSCAT 许可，仅行为定义，零代码行）——道莅 clean-room 实现
// 单位表：T[摄氏度] / Tw[摄氏度] / RH[%] / p[Pa] / p_ws[Pa] / e[Pa] /
//         gamma·p[Pa每摄氏度]
// 错误码表：16#0002_2F01 信息级（温度/湿度域外已钳位照算，或数值解超
//           承诺域下限被钳回 [摄氏度负 20]，不置 bError）/
//           16#0002_2F02 信息级（迭代达 40 次上限仍未达 0.05 摄氏度
//           区间精度，降级输出区间中点值，不置 bError——经验式本身是
//           近似）/ 16#0002_2F10 故障级（大气压非法或任一输入非有限，
//           置 bError）/ 16#0002_2F11 故障级（输入致二分区间非法：下界
//           残差非负、或终值自洽复检超容差，置 bError——该场景不可由
//           2F10 的输入幅值类判据观测，属区间构造独立域）/
//           16#0002_2F12 预留禁用（不得挪用）
// 状态机：N/A（纯函数；二分在单次调用内完成，无跨拍状态）
// 边界行为：① 干球温度域外（负 20~60 摄氏度外）钳位照算 + 信息 2F01，
//           头注释声明精度承诺收窄至负 20~60 摄氏度（Magnus 过水公式
//           拟合域外误差不承诺）；② RH 域外钳 1~100 + 信息 2F01；
//           ③ 大气压域外（50000~110000 Pa 外）→ 故障 2F10（v1.1.0
//           收窄声明：低压组合会使下界残差失去负号证明，见收敛域声明）；
//           ④ 二分 40 次未达精度 → 输出区间中点 + bValid := TRUE +
//           信息 2F02（降级可观测，不置故障）；⑤ 区间非法或自洽复检
//           失败 → 故障 2F11、bValid := FALSE、输出 0；异常路径输出
//           确定值，绝不输出未初始化值。
// 收敛域声明（R108 判据）：输入子域 T[负 20, 60] 摄氏度、RH[1, 100]%、
//           p[50000, 110000] Pa。收敛性论证：g(Tw) 在 Tw 上严格单调递增
//           （导数 = dp_ws/dTw + gamma·p > 0，过水 Magnus 斜率域内恒正）；
//           上界 g(T) = (1 - RH/100)·p_ws(T) >= 0（RH 钳后 <= 100 保证）；
//           下界 g(负 40) <= 19.0 - 0.000662·50000·20 - 1.04 < 0（取
//           p_ws(负 40) = 19.0 Pa、p >= 50000 Pa、T >= 负 20、RH >= 1
//           的最坏组合），故根必落于区间内，二分对区间宽度指数收敛，
//           无发散路径；低压域外（p < 50000）下界残差负号不再有保证，
//           按故障 2F10 拒绝而非静默外推。
// 验收向量推演（算法已证，手算，允差 ±0.1 摄氏度）：① T=30 摄氏度、
//           RH=65%、p=101325 Pa → Tw 约 24.8 摄氏度；② T=5 摄氏度、
//           RH=80%、p=101325 Pa → Tw 约 3.6 摄氏度；③ T=负 10 摄氏度、
//           RH=20%、p=101325 Pa → Tw 约 负 12.6 摄氏度；④ RH=100% 退化
//           → Tw = T 精确（g(T) = 0，区间上界即根）。编译器已证
//           （三平台）：未跑，由收口方登记。
// 修订历史：v1.0.0 2026-11-17 首版（R23 派单 · T1-2 焓湿图族拆分③ · 迭代式按检索原文修正）
//           v1.0.1 2026-11-17 R23 终审挂账警示（逻辑零改动）：DL_WB_GAMMA
//           1000 倍量纲错位 + 定点迭代在 e_s'(Tw)/(gamma·p) > 1 区间
//           结构性发散，修复前禁止用于生产数据链。
//           v1.1.0 2026-11-17 R24 挂账修复：二分法重写，引脚契约不变
//           （fTempC/fRh/fPress → fWetBulbC/bClamped/eErr/bError/bValid），
//           码位 2F01/2F02/2F10/2F11/2F12 全保留，语义重映射：2F02 =
//           迭代达上限未达 0.05 K 精度、2F11 = 输入致二分区间非法；
//           饱和压改 Magnus-Tetens 内联自洽实现，解除族属主件依赖。
//==============================================================================

FUNCTION FC_DL_WetBulbTempCalc : BOOL
VAR_INPUT
    fTempC  : LREAL;                     // 干球温度 [摄氏度]，有效域 -20.0..60.0，域外钳位照算 / Dry-bulb temperature [degC], valid range -20.0..60.0
    fRh     : LREAL;                     // 相对湿度 [百分数]，有效域 1.0..100.0，域外钳位照算 / Relative humidity [percent], valid range 1.0..100.0
    fPress  : LREAL := 101325.0;         // 大气压 [Pa]，有效域 50000..110000，域外故障拒绝 / Atmospheric pressure [Pa], valid range 50000..110000
END_VAR
VAR_OUTPUT
    fWetBulbC : LREAL;                   // 湿球温度 [摄氏度] / Wet-bulb temperature [degC]
    bClamped  : BOOL;                    // TRUE = 温度或湿度输入已钳位 / TRUE = temperature or humidity input clamped
    eErr      : UDINT;                   // 错误码，0 = 无错，码位 16#0002_2F01 起信息级、16#0002_2F10 起故障级（分带见错误码表） / Error code, 0 = no error, band info/fault per the code table
    bError    : BOOL;                    // 故障级标志，仅故障级错误置位 / Fault-class flag, set only on fault-level codes
    bValid    : BOOL;                    // 输出可用标志 / Outputs usable flag
END_VAR
VAR CONSTANT
    DL_WB_TMIN     : LREAL := -20.0;     // 承诺域下限 [摄氏度]，域外精度不承诺 / Promised domain floor [degC], accuracy not promised outside
    DL_WB_TMAX     : LREAL := 60.0;      // 承诺域上限 [摄氏度] / Promised domain ceiling [degC]
    DL_WB_BRACKET  : LREAL := -40.0;     // 二分区间下界 [摄氏度]，收敛域声明内恒有负残差 / Bisection bracket floor [degC]
    DL_WB_RH_MIN   : LREAL := 1.0;       // 湿度钳位下限 [百分数] / Humidity clamp floor [percent]
    DL_WB_RH_MAX   : LREAL := 100.0;     // 湿度钳位上限 [百分数] / Humidity clamp ceiling [percent]
    DL_WB_PMIN     : LREAL := 50000.0;   // 大气压有效域下限 [Pa] / Pressure domain floor [Pa]
    DL_WB_PMAX     : LREAL := 110000.0;  // 大气压有效域上限 [Pa] / Pressure domain ceiling [Pa]
    DL_WB_ITER_MAX : UINT  := 40;        // 二分迭代上限 [次]，防死锁计数器强制 / Bisection iteration ceiling [count], forced deadlock guard
    DL_WB_PREC     : LREAL := 0.05;      // 收敛精度：区间半宽 [摄氏度] / Convergence precision: bracket half-width [degC]
    DL_WB_GAMMA    : LREAL := 0.000662;  // 心理测量常数 gamma [1/摄氏度]（v1.1.0 量纲已修正） / Psychrometric constant gamma [1/degC], dimension fixed in v1.1.0
    DL_WB_MAGNUS_A : LREAL := 610.94;    // Magnus-Tetens 系数 A [Pa] / Magnus-Tetens coefficient A [Pa]
    DL_WB_MAGNUS_B : LREAL := 17.625;    // Magnus-Tetens 系数 B [无量纲] / Magnus-Tetens coefficient B [dimensionless]
    DL_WB_MAGNUS_C : LREAL := 243.04;    // Magnus-Tetens 系数 C [摄氏度] / Magnus-Tetens coefficient C [degC]
    DL_WB_RES_TOL  : LREAL := 50.0;      // 终值自洽复检容差 [Pa]（0.05 摄氏度区间对应残差带的上界） / Final residual recheck tolerance [Pa]
    DL_WB_EPS      : LREAL := 1.0E-6;    // 浮点判零容差 [混合] / Float zero tolerance
    DL_WB_INF      : LREAL := 1.7976931348623157E308; // LREAL 幅值上限 / LREAL magnitude ceiling
END_VAR
VAR
    fTEff    : LREAL;                    // 钳位后的生效干球温度 [摄氏度] / Effective clamped dry-bulb temperature [degC]
    fRhEff   : LREAL;                    // 钳位后的生效湿度 [百分数] / Effective clamped humidity [percent]
    fPwsT    : LREAL;                    // 干球温度下饱和压 p_ws(T) [Pa] / Saturation pressure at T [Pa]
    fVpAct   : LREAL;                    // 实际水汽压 e = RH/100·p_ws(T) [Pa] / Actual vapor pressure e [Pa]
    fGamPa   : LREAL;                    // 心理测量系数 gamma·p [Pa每摄氏度]，量纲已修正 / Psychrometric coefficient gamma times p [Pa/degC]
    fLo      : LREAL;                    // 二分区间下界 [摄氏度] / Bisection bracket low [degC]
    fHi      : LREAL;                    // 二分区间上界 [摄氏度] / Bisection bracket high [degC]
    fMid     : LREAL;                    // 二分中点 [摄氏度] / Bisection midpoint [degC]
    fResLo   : LREAL;                    // 下界残差 g(fLo) [Pa] / Bracket-low residual [Pa]
    fResMid  : LREAL;                    // 中点残差 g(fMid) [Pa] / Midpoint residual [Pa]
    fResFin  : LREAL;                    // 终值自洽复检残差 [Pa] / Final residual recheck [Pa]
    fMagDen  : LREAL;                    // Magnus 分母 (T + 243.04) [摄氏度] / Magnus denominator [degC]
    uIter    : UINT;                     // 迭代计数 [次] / Iteration counter [count]
END_VAR

(*------------------------------------------------------------------------------
 * 段 1｜出口默认值：入口即赋确定值
 *      Exit defaults: outputs assigned deterministically on entry
 *-----------------------------------------------------------------------------*)
FC_DL_WetBulbTempCalc := FALSE;          // 返回值默认无效 / Return value preset invalid
fWetBulbC := 0.0;                        // 湿球默认置零 / Wet bulb preset to zero
bClamped := FALSE;                       // 钳位标志默认 FALSE / Clamped flag preset FALSE
eErr := 16#0000_0000;                    // 错误码先清零 / Error code cleared first
bError := FALSE;                         // 故障标志先清零 / Fault flag cleared first
bValid := FALSE;                         // 可用标志先清零 / Usable flag cleared first

(*------------------------------------------------------------------------------
 * 段 2｜非有限值与大气压域闸门（R79 双侧幅值判 + v1.1.0 收窄域）
 *      Non-finite defense and the narrowed pressure-domain gate
 *-----------------------------------------------------------------------------*)
IF (fTempC <> fTempC) OR (ABS(fTempC) > DL_WB_INF)
   OR (fRh <> fRh) OR (ABS(fRh) > DL_WB_INF)
   OR (fPress <> fPress) OR (ABS(fPress) > DL_WB_INF) THEN
    eErr   := 16#0002_2F10;              // 故障级：输入非有限 / Fault: non-finite input
    bError := TRUE;                      // 置故障标志（R45 配对） / Raise the fault flag
    bValid := FALSE;                     // 输出不可用 / Outputs unusable
    RETURN;
END_IF
IF (fPress < DL_WB_PMIN) OR (fPress > DL_WB_PMAX) THEN
    eErr   := 16#0002_2F10;              // 故障级：大气压域外（收敛域声明外无负残差保证） / Fault: pressure outside the convergence domain
    bError := TRUE;                      // 置故障标志 / Raise the fault flag
    bValid := FALSE;                     // 输出不可用 / Outputs unusable
    RETURN;
END_IF

(*------------------------------------------------------------------------------
 * 段 3｜输入钳位：温度 -20~60、湿度 1~100，信息级共码 2F01（R90）
 *      Input clamping, shared info code per R90
 *-----------------------------------------------------------------------------*)
IF (fTempC < DL_WB_TMIN) OR (fTempC > DL_WB_TMAX) THEN
    fTEff := MIN(MAX(fTempC, DL_WB_TMIN), DL_WB_TMAX); // 温度双侧钳位 / Two-sided temperature clamp
    bClamped := TRUE;                    // 钳位声明置位 / Clamped flag raised
    eErr := 16#0002_2F01;                // 信息级：输入已钳位（不置 bError） / Info: input clamped, no fault flag
ELSE
    fTEff := fTempC;                     // 合法温度原值生效 / Valid temperature applied as-is
END_IF
IF (fRh < DL_WB_RH_MIN) OR (fRh > DL_WB_RH_MAX) THEN
    fRhEff := MIN(MAX(fRh, DL_WB_RH_MIN), DL_WB_RH_MAX); // 湿度双侧钳位 / Two-sided humidity clamp
    bClamped := TRUE;                    // 钳位声明置位 / Clamped flag raised
    eErr := 16#0002_2F01;                // 信息级：输入已钳位 / Info: input clamped
ELSE
    fRhEff := fRh;                       // 合法湿度原值生效 / Valid humidity applied as-is
END_IF

(*------------------------------------------------------------------------------
 * 段 4｜系数与残差量预置：Magnus-Tetens 内联（与残差同源自洽）
 *      Coefficients preset, Magnus-Tetens inline, self-consistent
 *-----------------------------------------------------------------------------*)
fMagDen := fTEff + DL_WB_MAGNUS_C;       // Magnus 分母 [摄氏度]，域内恒 >= 203 / Magnus denominator, always >= 203 in domain
IF fMagDen <= DL_WB_EPS THEN
    eErr   := 16#0002_2F11;              // 故障级：分母退化归区间非法（域内不可达，防御兜底） / Fault: degenerate denominator folded into the bracket fault
    bError := TRUE;                      // 置故障标志 / Raise the fault flag
    bValid := FALSE;                     // 输出不可用 / Outputs unusable
    RETURN;
END_IF
fPwsT  := DL_WB_MAGNUS_A * EXP(DL_WB_MAGNUS_B * fTEff / fMagDen); // 干球饱和压 [Pa] / Saturation pressure at T [Pa]
fVpAct := (fRhEff / 100.0) * fPwsT;      // 实际水汽压 e [Pa] / Actual vapor pressure e [Pa]
fGamPa := DL_WB_GAMMA * fPress;          // 心理测量系数 gamma·p [Pa每摄氏度] / Psychrometric coefficient [Pa/degC]

(*------------------------------------------------------------------------------
 * 段 5｜区间构造与合法性闸：g 单调增，要求 g(fLo) < 0 <= g(fHi)
 *      Bracket construction and validity gate
 *-----------------------------------------------------------------------------*)
fLo := DL_WB_BRACKET;                    // 下界 -40 摄氏度 / Bracket low
fHi := fTEff;                            // 上界取干球 / Bracket high, the dry bulb
fResLo := DL_WB_MAGNUS_A * EXP(DL_WB_MAGNUS_B * fLo / (fLo + DL_WB_MAGNUS_C))
          - fGamPa * (fTEff - fLo) - fVpAct; // 下界残差 g(fLo) [Pa] / Bracket-low residual [Pa]
IF fResLo >= DL_WB_EPS THEN
    fWetBulbC := 0.0;                    // 区间非法：丢弃结果 / Illegal bracket, result discarded
    eErr   := 16#0002_2F11;              // 故障级：输入致二分区间非法 / Fault: input-induced illegal bracket
    bError := TRUE;                      // 置故障标志 / Raise the fault flag
    bValid := FALSE;                     // 输出不可用 / Outputs unusable
    RETURN;
END_IF

(*------------------------------------------------------------------------------
 * 段 6｜二分迭代：区间半宽收敛于 0.05 摄氏度，计数器强制防死锁
 *      Bisection loop, counter-forced deadlock guard
 *-----------------------------------------------------------------------------*)
uIter := 0;                              // 迭代计数清零 / Counter cleared
WHILE ((fHi - fLo) > DL_WB_PREC) AND (uIter < DL_WB_ITER_MAX) DO
    fMid := 0.5 * (fLo + fHi);           // 区间中点 [摄氏度] / Bracket midpoint
    fMagDen := fMid + DL_WB_MAGNUS_C;    // Magnus 分母 [摄氏度] / Magnus denominator
    IF fMagDen <= DL_WB_EPS THEN
        fWetBulbC := 0.0;                // 分母退化：丢弃结果 / Degenerate denominator, result discarded
        eErr   := 16#0002_2F11;          // 故障级：退化归区间非法（R90） / Fault: degeneracy folded into the bracket fault
        bError := TRUE;                  // 置故障标志 / Raise the fault flag
        bValid := FALSE;                 // 输出不可用 / Outputs unusable
        RETURN;
    END_IF
    fResMid := DL_WB_MAGNUS_A * EXP(DL_WB_MAGNUS_B * fMid / fMagDen)
               - fGamPa * (fTEff - fMid) - fVpAct; // 中点残差 g(fMid) [Pa] / Midpoint residual [Pa]
    IF fResMid >= 0.0 THEN
        fHi := fMid;                     // 根在中点以下，上界下压 / Root below midpoint, lower the high bound
    ELSE
        fLo := fMid;                     // 根在中点以上，下界上抬 / Root above midpoint, raise the low bound
    END_IF
    uIter := uIter + 1;                  // 计数递增（防死锁强制项） / Counter increment, the forced guard
END_WHILE
fMid := 0.5 * (fLo + fHi);               // 终值取区间中点 / Final value is the bracket midpoint

(*------------------------------------------------------------------------------
 * 段 7｜终值自洽复检与输出域钳回：残差超容差归 2F11；越 -20 钳回 + 2F01
 *      Final residual recheck and output-domain clamp
 *-----------------------------------------------------------------------------*)
fMagDen := fMid + DL_WB_MAGNUS_C;        // Magnus 分母 [摄氏度] / Magnus denominator
IF fMagDen <= DL_WB_EPS THEN
    fWetBulbC := 0.0;                    // 退化：丢弃结果 / Degenerate, result discarded
    eErr   := 16#0002_2F11;              // 故障级：退化归区间非法（R90） / Fault: degeneracy folded into the bracket fault
    bError := TRUE;                      // 置故障标志 / Raise the fault flag
    bValid := FALSE;                     // 输出不可用 / Outputs unusable
    RETURN;
END_IF
fResFin := DL_WB_MAGNUS_A * EXP(DL_WB_MAGNUS_B * fMid / fMagDen)
           - fGamPa * (fTEff - fMid) - fVpAct; // 终值残差 [Pa] / Final residual [Pa]
IF ABS(fResFin) > DL_WB_RES_TOL THEN
    fWetBulbC := 0.0;                    // 自洽复检失败：丢弃结果 / Self-consistency failed, result discarded
    eErr   := 16#0002_2F11;              // 故障级：复检失败归区间非法语义（R90） / Fault: recheck failure folded into the bracket fault
    bError := TRUE;                      // 置故障标志 / Raise the fault flag
    bValid := FALSE;                     // 输出不可用 / Outputs unusable
    RETURN;
END_IF
IF fMid < DL_WB_TMIN THEN
    fMid := DL_WB_TMIN;                  // 数值解越承诺域下限，钳回 -20 / Numerical solution below the promised floor, clamped back
    eErr := 16#0002_2F01;                // 信息级：解域下限钳回（不置 bError） / Info: solution clamped to the floor, no fault flag
END_IF
IF fMid > fTEff THEN
    fMid := fTEff;                       // 数值上溢钳回干球（湿球不超过干球） / Numerical overshoot clamped to the dry bulb
END_IF
fWetBulbC := fMid;                       // 湿球温度出口 / Wet-bulb temperature outlet
IF uIter >= DL_WB_ITER_MAX THEN
    eErr := 16#0002_2F02;                // 信息级：40 次未达精度，降级输出中点（不置故障） / Info: iteration ceiling met without precision, degraded midpoint, no fault
END_IF
bValid := TRUE;                          // 输出可用（含降级情形，见 2F02 口径） / Outputs usable, including the degraded case
FC_DL_WetBulbTempCalc := TRUE;           // 返回 TRUE = 计算有效 / Return TRUE = computation valid
END_FUNCTION

(* ---- FC_DL_WrapToRange.st ---- *)
(*==============================================================================
 * 名称 : FC_DL_WrapToRange —— 周期量卷绕到 [fLo,fHi)（区间宽度 <=0 判参数非法）
 * 分类 / 前缀 / 版本 : DL_Algo / FC_DL_ / 1.0.0
 * 溯源 : 开源语义参考（OSCAT/AixOCAT 族，MIT）或 clean-room IEC 实现，未复制源码
 * 平台 : 纯 IEC 61131-3
 * 功能说明 : 将任意输入卷绕到 [fLo, fHi) 周期区间：先平移到以 fLo 为原点，
 *            整周期 TRUNC 截断缩圈，负余量加一周期修正，再加回 fLo。
 *            例：区间 [0,360)、输入 -10 → 350；区间 [100,200)、输入 250 → 150。
 *            边界处理：fHi-fLo<=0 判参数非法（防除零，区间无宽度）；任一
 *            输入非有限（NaN/±Inf）置 eErr 返回 0.0；TRUNC 为 LREAL 通用
 *            形式无整型溢出，结果落在 [fLo,fHi) 左闭右开。
 * 错误码 : 16#0001_1C06 = 区间宽度非法（fHi<=fLo），或输入非有限（NaN/±Inf）
 *          eErr=0 且 bValid=TRUE 表示卷绕结果可用
 * 状态机 : R6 标注 N/A（纯函数无顺序状态，以本节替代 ELSE 兜底）
 * 红线 : R1/R2/R3 ✓ 零全局/零IO/纯IEC ｜ R4 ✓ 非有限拦截/除零防护（宽度校验）｜ R10 ✓ 标准转换 ｜ R11 ✓ 分号收尾 ｜ R15 ✓ 无保留字撞名
 * 修订记录 : 2026-11-23 v1.0.0 首次入库（R76）
 *============================================================================*)
FUNCTION FC_DL_WrapToRange : LREAL
VAR_INPUT
    fIn : LREAL;    // 待卷绕输入量 [工程单位] / input value to wrap
    fLo : LREAL;    // 区间下界（含）[工程单位] / range lower bound, inclusive
    fHi : LREAL;    // 区间上界（不含）[工程单位] / range upper bound, exclusive
END_VAR
VAR_OUTPUT
    eErr   : UDINT;    // 故障码，0=正常，1C06=区间非法或非有限 / error code
    bError : BOOL;     // TRUE=本件发生故障 / TRUE when fault occurred
    bValid : BOOL;     // TRUE=卷绕结果可用 / TRUE when result is usable
END_VAR
VAR
    _fW : LREAL;       // 区间宽度（周期）[工程单位] / range width as period
    _fR : LREAL;       // 平移后的余量 [工程单位] / offset remainder
END_VAR

FC_DL_WrapToRange := 0.0;                    // 返回值预设 0.0 / preset return to zero
eErr   := 16#0000_0000;                      // 故障码清零 / clear error code
bError := FALSE;                             // 故障标志清零 / clear error flag
bValid := TRUE;                              // 预设输出可用 / preset valid flag

IF (fIn <> fIn) OR ((fIn - fIn) <> (fIn - fIn))          // fIn 非有限 / NaN or infinite
   OR (fLo <> fLo) OR ((fLo - fLo) <> (fLo - fLo))        // fLo 非有限 / NaN or infinite
   OR (fHi <> fHi) OR ((fHi - fHi) <> (fHi - fHi)) THEN   // fHi 非有限 / NaN or infinite
    eErr   := 16#0001_1C06;                  // 置非有限故障码 / set non-finite code
    bError := TRUE;                          // 置故障标志 / set error flag
    bValid := FALSE;                         // 输出不可用 / outputs not usable
    RETURN;                                  // 返回 0.0 / return zero
END_IF

_fW := fHi - fLo;                            // 计算区间宽度 / compute range width
IF _fW <= 0.0 THEN                           // 宽度非正：参数非法且防除零 / non-positive width invalid
    eErr   := 16#0001_1C06;                  // 置区间非法码 / set invalid-range code
    bError := TRUE;                          // 置故障标志 / set error flag
    bValid := FALSE;                         // 输出不可用 / outputs not usable
    RETURN;                                  // 返回 0.0 / return zero
END_IF

_fR := fIn - fLo;                            // 平移到原点 / shift origin to fLo
_fR := _fR - _fW * TRUNC(_fR / _fW);         // 整周期截断缩圈（TRUNC 向零，防除零已保证）/ strip whole periods
IF _fR < 0.0 THEN                            // 负余量修正 / fix negative remainder
    _fR := _fR + _fW;                        // 加一周期 / add one period
END_IF

FC_DL_WrapToRange := fLo + _fR;              // 加回下界，落 [fLo,fHi) / restore origin

END_FUNCTION

(* ---- FB_DL_AdaptiveDeadbandZone.st ---- *)
(*
  Name        : FB_DL_AdaptiveDeadbandZone
  Category    : DL_Algo
  Version     : 1.0.0
  Purpose     : 噪声带自适应死区：以一阶差分绝对值的 EMA 在线估计噪声幅值，按倍率整定死区宽度（上下限可组态），输出死区后信号仅供显示/滤波链使用；/ Noise-adaptive deadband: estimate noise amplitude by EMA of absolute first differences, scale it into a configurable deadband width, output the deadbanded signal
  溯源        : 借 t2-5-modpid·deadband 的分类/参数域组织，clean-room 实现
  Boundary    : ① 组态闸：fDbMax - fDbMin <= eps / fDbMin < 0 / fNoiseGain <= 0 / fAlpha 不在 (0,1] → 锁存故障，输出保持；
                ② 非有限输入该拍不更新噪声估计与输出（保留上拍值）；
                ③ 死区判据 |fIn - fOut| > db 用容差比较（禁 = / <>）；
                ④ 首拍无前值时以当前输入初始化，不产生虚假大差分（隐性回夹防护）；
                ⑤ 倍率钳位：db 先按 [fDbMin, fDbMax] 饱和再参与判据，饱和方向为「更保守的大死区」。
*)
TYPE E_DL_AdzState :
(
    eIdle  := 0,                             (* 未使能 / Disabled *)
    eRun   := 10,                            (* 自适应运行 / Adaptive running *)
    eFault := 90                             (* 故障锁存相 / Fault latched *)
);
END_TYPE

TYPE E_DL_AdzCause :
(
    eNone       := 0,                        (* 无故障成因 / No cause *)
    eCfgIllegal := 1,                        (* 组态非法：限值/倍率/系数越域 / Illegal config *)
    ePhaseBad   := 2                         (* 非法相位兜底 / Illegal phase fallback *)
);
END_TYPE

FUNCTION_BLOCK FB_DL_AdaptiveDeadbandZone
VAR_INPUT
    fIn        : REAL := 0.0;                (* 原始测量输入（噪声信号）[工程单位] / Raw noisy measurement *)
    fNoiseGain : REAL := 3.0;                (* 噪声→死区倍率（典型 2..4），域 > 0 [-] / Noise to deadband gain, > 0 *)
    fDbMin     : REAL := 0.0;                (* 死区下限，域 >= 0 [工程单位] / Deadband lower limit, >= 0 *)
    fDbMax     : REAL := 10.0;               (* 死区上限，域 > fDbMin [工程单位] / Deadband upper limit *)
    fAlpha     : REAL := 0.2;                (* 噪声 EMA 新值权重，域 (0, 1] [-] / Noise EMA weight, (0,1] *)
    bEnable    : BOOL := TRUE;               (* 使能 [-] / Enable *)
    bReset     : BOOL := FALSE;              (* 复位命令，上升沿清噪声估计与输出 [-] / Reset command *)
END_VAR
VAR_OUTPUT
    fOut       : REAL;                       (* 死区处理后信号 [工程单位] / Deadbanded signal *)
    fDeadband  : REAL;                       (* 当前生效死区宽度（半宽）[工程单位] / Effective deadband half-width *)
    fNoiseEst  : REAL;                       (* 噪声幅值估计（|Δ| EMA）[工程单位] / Estimated noise amplitude *)
    bDbActive  : BOOL;                       (* 死区正在吞掉变化（本拍输出保持）[-] / Deadband currently suppressing *)
    eState     : E_DL_AdzState;              (* 状态出口 / State outlet *)
    eCause     : E_DL_AdzCause;              (* 故障成因出口（R190 归因唯一） / Fault cause outlet *)
    bError     : BOOL;                       (* 故障锁存标志 [-] / Fault latch flag *)
END_VAR
VAR
    _eState   : E_DL_AdzState := E_DL_AdzState.eIdle;    (* 内部相位（CASE 唯一写入目标） / Internal phase *)
    _eCause   : E_DL_AdzCause := E_DL_AdzCause.eNone;    (* 故障成因锁存量 / Latched cause *)
    rtReset   : R_TRIG;                      (* 复位沿实例，段 0 无条件调用 / Reset edge instance *)
    _bFault   : BOOL;                        (* 故障锁存位 / Latched fault bit *)
    _bCfgBad  : BOOL;                        (* 组态非法当拍量 / Illegal config this scan *)
    _bInit    : BOOL;                        (* 前值初始化标志（首拍不产虚假差分） / First-scan init flag *)
    _bFinite  : BOOL;                        (* 输入有限性当拍量 / Input finiteness this scan *)
    _fPrev    : REAL;                        (* 上拍输入快照（差分基准）[工程单位] / Previous input snapshot *)
    _fDiff    : REAL;                        (* 本拍一阶差分绝对值 [工程单位] / Absolute first difference *)
    _fNoise   : REAL;                        (* 噪声幅值 EMA 内部量 [工程单位] / Noise EMA internal *)
    _fDb      : REAL;                        (* 未钳位死区 = 倍率 × 噪声 [工程单位] / Unclamped deadband *)
    _fDelta   : REAL;                        (* |输入 - 输出| 偏离量（判据用）[工程单位] / Deviation magnitude *)
    _fOne     : REAL;                        (* 实数 1 常量（EMA 系数补数用）[-] / Real one constant *)
END_VAR
VAR CONSTANT
    DL_ADZ_EPS : REAL := 1.0E-6;             (* 容差（REAL 量级，带宽/系数/比较共用）[-] / Tolerance epsilon *)
END_VAR

(* —— 段 0：当拍判据派生 + 实例无条件刷新（R228A） —— *)
_bCfgBad := ((fDbMax - fDbMin) <= DL_ADZ_EPS)                                  (* 死区上下限颠倒闸 / Band inversion gate *)
            OR (fDbMin < 0.0)                                                  (* 下限负域闸 / Negative lower-limit gate *)
            OR (fNoiseGain <= DL_ADZ_EPS)                                      (* 倍率正域闸（防死区恒 0 或取反） / Gain positive gate *)
            OR (fAlpha <= DL_ADZ_EPS) OR (fAlpha > 1.0);                       (* EMA 系数域闸 (0,1] / EMA weight gate *)
rtReset(CLK := bReset);                                                        (* 复位沿每拍必调 / Reset edge every scan *)
_bFinite := (fIn = fIn) AND ((fIn - fIn) = (fIn - fIn));                       (* NaN 自反 + Inf 差判联合闸 / NaN and Inf gate *)
_fOne := 1.0;                                                                  (* 常量装载（避免字面量散布） / Constant load *)

(* —— 段 1：单拍量预清零（R107） —— *)
bDbActive := FALSE;                                                            (* 死区抑制指示预清 / Suppression preset *)

(* —— 段 2：复位沿处理（作用域：清故障 + 清噪声估计 + 清初始化 + 迁 eIdle，R283 逐项声明） —— *)
IF rtReset.Q THEN
    _bFault := FALSE;                                                          (* 清故障锁存 / Clear fault *)
    _eCause := E_DL_AdzCause.eNone;                                            (* 清成因 / Clear cause *)
    _fNoise := 0.0;                                                            (* 清噪声估计 / Clear noise estimate *)
    _fPrev := 0.0;                                                             (* 清差分基准 / Clear previous sample *)
    _bInit := FALSE;                                                           (* 清初始化标志（首拍重新对齐） / Clear init flag *)
    fOut := 0.0;                                                               (* 清输出 / Clear output *)
    fDeadband := fDbMin;                                                       (* 死区回下限（组态基准值） / Deadband back to lower limit *)
    fNoiseEst := 0.0;                                                          (* 清噪声出口 / Clear noise outlet *)
    _eState := E_DL_AdzState.eIdle;                                            (* 迁未使能相 / Back to idle *)
END_IF

(* —— 段 3：组态故障锁存（锁存至复位沿，R189） —— *)
IF _bCfgBad AND NOT _bFault THEN
    _bFault := TRUE;                                                           (* 锁存故障位 / Latch fault *)
    _eCause := E_DL_AdzCause.eCfgIllegal;                                      (* 成因：组态非法 / Cause: illegal config *)
    _eState := E_DL_AdzState.eFault;                                           (* 同步迁故障相 / Migrate to fault *)
END_IF

(* —— 段 4：CASE 主状态机（ELSE 兜底迁 eFault，红线 6） —— *)
CASE _eState OF
    E_DL_AdzState.eIdle:                                                       (* 未使能：输出直通、死区置下限 / Disabled *)
        _bInit := FALSE;                                                       (* 失能清初始化，重使能时重新对齐 / Clear init while disabled *)
        fDeadband := fDbMin;                                                   (* 死区取组态下限 / Deadband = lower limit *)
        IF bEnable AND NOT _bFault THEN
            _eState := E_DL_AdzState.eRun;                                     (* 使能进入自适应 / Enter adaptive *)
        END_IF
    E_DL_AdzState.eRun:                                                        (* 自适应相：噪声估计 + 死区整定 + 死区输出 / Adaptive *)
        IF NOT bEnable THEN
            _eState := E_DL_AdzState.eIdle;                                    (* 失能回未使能 / Back to idle *)
        ELSIF _bFinite THEN
            IF NOT _bInit THEN
                _fPrev := fIn;                                                 (* 首拍对齐：基准取当前输入（防虚假大差分） / First scan alignment *)
                fOut := fIn;                                                   (* 首拍直通（无历史可比） / First scan passthrough *)
                _bInit := TRUE;                                                (* 立初始化标志 / Set init flag *)
            END_IF
            _fDiff := ABS(fIn - _fPrev);                                       (* 一阶差分绝对值（噪声代理）[工程单位] / Absolute first difference *)
            _fNoise := (1.0 - fAlpha) * _fNoise + fAlpha * _fDiff;             (* 噪声 EMA（系数和恒 1，无漂移） / Noise EMA *)
            _fPrev := fIn;                                                     (* 快照推进（仅有限拍推进） / Advance snapshot *)
            _fDb := fNoiseGain * _fNoise;                                      (* 倍率映射到死区半宽 / Gain to deadband *)
            IF _fDb < fDbMin THEN
                _fDb := fDbMin;                                                (* 下限饱和：死区不小于组态下限 / Lower saturation *)
            ELSIF _fDb > fDbMax THEN
                _fDb := fDbMax;                                                (* 上限饱和：防死区吞掉真实变化过大 / Upper saturation *)
            END_IF
            fDeadband := _fDb;                                                 (* 死区出口（实时派生） / Deadband outlet *)
            fNoiseEst := _fNoise;                                              (* 噪声估计出口 / Noise outlet *)
            _fDelta := ABS(fIn - fOut);                                        (* 与当前输出的偏离量 / Deviation from output *)
            IF _fDelta > _fDb THEN
                fOut := fIn;                                                   (* 偏离超死区：输出跟随（更新） / Exceeds band: follow *)
                bDbActive := FALSE;                                            (* 未抑制 / Not suppressing *)
            ELSE
                bDbActive := TRUE;                                             (* 偏离在带内：输出保持（抑制噪声） / Within band: hold *)
            END_IF
        END_IF                                                                 (* 非有限输入：噪声估计与输出均保持上拍（边界②） / Non-finite: hold *)
    E_DL_AdzState.eFault:                                                      (* 故障相：冻结保持末值，仅复位沿出 / Fault *)
        ;                                                                      (* 锁存回放（R28） / Replay from latch *)
    ELSE                                                                       (* 非法相位兜底迁安全态 / Illegal phase fallback *)
        _eState := E_DL_AdzState.eFault;                                       (* 迁故障相 / To fault *)
        _bFault := TRUE;                                                       (* 同步锁存 / Latch *)
        _eCause := E_DL_AdzCause.ePhaseBad;                                    (* 成因：非法相位 / Cause: illegal phase *)
END_CASE

(* —— 段 5：出口映射（bError/eState 同源，R191） —— *)
bError := _bFault;                                                             (* 故障标志镜像 / Fault flag mirror *)
eState := _eState;                                                             (* 状态出口 / State outlet *)
eCause := _eCause;                                                             (* 成因出口 / Cause outlet *)
END_FUNCTION_BLOCK
